TYPE ST_EL3312ChannelState_1 :
STRUCT
	bUnderrange				:BOOL;			(* State underrange *)
	bOverrange				:BOOL;			(* State overrange *)
	byLimit1					:BYTE;			(* State limit 1 *)
	byLimit2 					:BYTE;			(* State limit 2 *)
	bError 					:BOOL;			(* State error *)
	bState 					:BOOL;			(* State *)
	bToggle					:BOOL;			(* TxPDO Toggle *)
END_STRUCT
END_TYPE

(* stored: Version 1.1.0.1, ProductVersion 3.1.4024.15
   DUT ST_EL3312ChannelState_1: Id {3d8048a0-f03c-4275-9b69-4bbfc4d10c7b} *)
